TYPE "FRK_ProbeRow"
VERSION : 0.1
STRUCT
    BeginCalls : DInt;
    EndCalls : DInt;
    InitCalls : DInt;
    CyclicCalls : DInt;
    BeginOrder : DInt;
    InitOrder : DInt;
END_STRUCT;
END_TYPE
